(* IEC 61131-3 sources: plc-vscode/tests/st/all/rusty/tests/lit/multi/cross_unit_struct_init, 2 files *)

(* ---- main.st ---- *)
// CHECK: 42
// CHECK: 10

TYPE MyStruct : STRUCT
    fb : FbA;
    v  : myINT;
END_STRUCT
END_TYPE

FUNCTION main : DINT
VAR
    s : MyStruct;
END_VAR
    printf('%d$N', s.fb.x);
    printf('%d$N', s.v);
END_FUNCTION

(* ---- fb_def.st ---- *)
FUNCTION_BLOCK FbA
VAR
    x : DINT := 42;
END_VAR
END_FUNCTION_BLOCK

TYPE myINT : INT := 10; END_TYPE
